(*
SPDX-FileCopyrightText: © 2026 Oleksandr Tiutyk <trofimich@gmail.com>
SPDX-License-Identifier: MIT
License: https://opensource.org/license/mit
*)

(*
Identifies the cyclic step of the auto-disposed object registry growth and reuse regression test.
*)
{attribute 'qualified_only'}
{attribute 'strict'}
{attribute 'to_string'}
TYPE DYNAMIC_MEMORY_REGISTRY_GROWTH_PHASE :
(
	REGISTER_GROWING_BATCH,
	VERIFY_GROWING_BATCH_AND_REUSE,
	VERIFY_REUSED_BATCH
);
END_TYPE

(* stored: Version 1.1.0.1, ProductVersion 3.1.4026.21
   DUT DYNAMIC_MEMORY_REGISTRY_GROWTH_PHASE: Id {83482883-1251-4ac3-bc1c-41ad87742585} *)
